(* IEC 61131-3 sources: stdmachine/plc/src/01_Types, 123 files *)

(* ---- E_ActStatus.st ---- *)
// Statut de l'action d'un objet (docs/04 § 5)
{attribute 'qualified_only'}
{attribute 'strict'}
TYPE E_ActStatus :
(
    Idle := 0,
    Busy := 1,
    Done := 2,
    Error := 3
) USINT;
END_TYPE

(* ---- E_AlarmEvent.st ---- *)
// Événement d'alarme (docs/14 § 5)
{attribute 'qualified_only'}
{attribute 'strict'}
TYPE E_AlarmEvent :
(
    Raised := 0,
    Cleared := 1,
    Acked := 2,
    Repeated := 3,
    Closed := 4
) USINT;
END_TYPE

(* ---- E_AlarmState.st ---- *)
// État d'une alarme active (docs/14 § 5)
{attribute 'qualified_only'}
{attribute 'strict'}
TYPE E_AlarmState :
(
    ActiveUnacked := 0,
    ActiveAcked := 1,
    ClearedUnacked := 2
) USINT;
END_TYPE

(* ---- E_BindTarget.st ---- *)
// Cible d'une liaison de résultat ou d'un SetVar (docs/06 § 2)
{attribute 'qualified_only'}
{attribute 'strict'}
TYPE E_BindTarget :
(
    None := 0,
    Var := 1,
    PartData := 2,
    PartId := 3,
    Verdict := 4,
    PartRemoved := 5,
    MoverData := 6,
    Output := 7
) USINT;
END_TYPE

(* ---- E_CalibState.st ---- *)
// État d'une calibration (docs/05 § 10.1)
{attribute 'qualified_only'}
{attribute 'strict'}
TYPE E_CalibState :
(
    Never := 0,
    Valid := 1,
    Expired := 2,
    Failed := 3,
    Running := 4
) USINT;
END_TYPE

(* ---- E_Cmd.st ---- *)
// Commandes d'état (docs/02 § 8). DrainStart et DrainCancel ne concernent que la machine (docs/05 § 5.7) :
// FB_PackML les ignore, le séquenceur général les traite.
{attribute 'qualified_only'}
{attribute 'strict'}
TYPE E_Cmd :
(
    None := 0,
    Reset := 1,
    Start := 2,
    Stop := 3,
    Hold := 4,
    Abort := 5,
    Clear := 6,
    DrainStart := 7,
    DrainCancel := 8
) USINT;
END_TYPE

(* ---- E_CmdResult.st ---- *)
// Résultat d'une commande (docs/05 § 2, docs/06 § 6.1)
{attribute 'qualified_only'}
{attribute 'strict'}
TYPE E_CmdResult :
(
    None := 0,
    Accepted := 1,
    Rejected := 2
) USINT;
END_TYPE

(* ---- E_Cmp.st ---- *)
// Comparaison d'un terme de condition (docs/05 § 3.7)
{attribute 'qualified_only'}
{attribute 'strict'}
TYPE E_Cmp :
(
    Eq := 0,
    Ne := 1,
    Lt := 2,
    Le := 3,
    Gt := 4,
    Ge := 5,
    IsTrue := 6,
    IsFalse := 7
) USINT;
END_TYPE

(* ---- E_Combine.st ---- *)
// Combinaison des termes d'une condition (docs/05 § 3.7)
{attribute 'qualified_only'}
{attribute 'strict'}
TYPE E_Combine :
(
    All := 0,
    Any := 1
) USINT;
END_TYPE

(* ---- E_CtxStatus.st ---- *)
// Statut d'un contexte d'exécution (docs/05 § 3.1)
{attribute 'qualified_only'}
{attribute 'strict'}
TYPE E_CtxStatus :
(
    Free := 0,
    Running := 1,
    WaitAction := 2,
    WaitCond := 3,
    WaitTime := 4,
    WaitJoin := 5,
    WaitStep := 6,
    Holding := 7,
    Done := 8,
    Failed := 9
) USINT;
END_TYPE

(* ---- E_DeclaredState.st ---- *)
// État déclaré de la machine (docs/12 § 2)
{attribute 'qualified_only'}
{attribute 'strict'}
TYPE E_DeclaredState :
(
    None := 0,
    PlannedStop := 1,
    Changeover := 2,
    WaitUpstream := 3,
    WaitDownstream := 4,
    PlannedMaintenance := 5,
    CorrectiveMaintenance := 6,
    Trials := 7,
    Cleaning := 8
) USINT;
END_TYPE

(* ---- E_DeployCmd.st ---- *)
// Commande de déploiement (docs/05 § 10)
{attribute 'qualified_only'}
{attribute 'strict'}
TYPE E_DeployCmd :
(
    None := 0,
    Verify := 1,
    Activate := 2,
    Cancel := 3
) USINT;
END_TYPE

(* ---- E_FailPolicy.st ---- *)
// Politique d'échec d'une instruction Action (docs/05 § 3.6)
{attribute 'qualified_only'}
{attribute 'strict'}
TYPE E_FailPolicy :
(
    StopStation := 0,
    Retry := 1,
    PartBad := 2,
    Goto := 3,
    Ignore := 4
) USINT;
END_TYPE

(* ---- E_ForceKind.st ---- *)
// Nature d'un forçage (docs/12 § 7)
{attribute 'qualified_only'}
{attribute 'strict'}
TYPE E_ForceKind :
(
    None := 0,
    DeclaredState := 1,
    StationOutOfProduction := 2,
    MoverOutOfService := 3
) USINT;
END_TYPE

(* ---- E_GroupRole.st ---- *)
// Rôle d'une fonction (docs/06 § 4)
{attribute 'qualified_only'}
{attribute 'strict'}
TYPE E_GroupRole :
(
    Entry := 0,
    Work := 1,
    Exit := 2,
    Reject := 3
) USINT;
END_TYPE

(* ---- E_Judgement.st ---- *)
// Jugement d'un résultat (docs/04 § 5)
{attribute 'qualified_only'}
{attribute 'strict'}
TYPE E_Judgement :
(
    None := 0,
    Ok := 1,
    Nok := 2,
    High := 3,
    Low := 4
) USINT;
END_TYPE

(* ---- E_ManualKind.st ---- *)
// Nature d'une demande du canal manuel (docs/05 § 7)
{attribute 'qualified_only'}
{attribute 'strict'}
TYPE E_ManualKind :
(
    Action := 0,
    JogStart := 1,
    JogStop := 2,
    Ack := 3,
    TeachPosition := 4
) USINT;
END_TYPE

(* ---- E_Mode.st ---- *)
// Modes de la machine (docs/02 § 8)
{attribute 'qualified_only'}
{attribute 'strict'}
TYPE E_Mode :
(
    Production := 0,
    Maintenance := 1
) USINT;
END_TYPE

(* ---- E_MoverState.st ---- *)
// État d'un mover dans le séquenceur général (docs/05 § 5.3)
{attribute 'qualified_only'}
{attribute 'strict'}
TYPE E_MoverState :
(
    Unknown := 0,
    Ready := 1,
    Routing := 2,
    Queued := 3,
    AtStation := 4,
    Buffered := 5,
    ToEmpty := 6,
    Error := 7,
    Halted := 8,
    OutOfService := 9
) USINT;
END_TYPE

(* ---- E_MoverVarReset.st ---- *)
// Règle de remise à zéro d'une variable de mover (docs/05 § 5.8)
{attribute 'qualified_only'}
{attribute 'strict'}
TYPE E_MoverVarReset :
(
    Never := 0,
    OnDeploy := 1,
    OnEmpty := 2
) USINT;
END_TYPE

(* ---- E_ObjState.st ---- *)
// États d'un objet (docs/04 § 5 et § 7.1)
{attribute 'qualified_only'}
{attribute 'strict'}
TYPE E_ObjState :
(
    NotInitialized := 0,
    Ready := 1,
    Busy := 2,
    Error := 3,
    Disabled := 4
) USINT;
END_TYPE

(* ---- E_Op.st ---- *)
// Jeu d'instructions (docs/06 § 2) ; version 2 du jeu : 17 à 23
{attribute 'qualified_only'}
{attribute 'strict'}
TYPE E_Op :
(
    Nop := 0,
    Action := 1,
    WaitCond := 2,
    WaitTime := 3,
    Jump := 4,
    JumpIfFalse := 5,
    Fork := 6,
    Join := 7,
    LoopInit := 8,
    LoopNext := 9,
    Call := 10,
    Return := 11,
    SetVar := 12,
    Alarm := 13,
    End := 14,
    StepBegin := 15,
    StepEnd := 16,
    WaitMover := 17,
    Prompt := 18,
    SavePos := 19,
    Route := 20,
    CalibStation := 21,
    ResetMoverVars := 22,
    SetOut := 23
) UINT;
END_TYPE

(* ---- E_OpStatus.st ---- *)
// Réponse d'une station à une demande d'opération (docs/05 § 4.1)
{attribute 'qualified_only'}
{attribute 'strict'}
TYPE E_OpStatus :
(
    Idle := 0,
    Running := 1,
    Done := 2,
    Failed := 3,
    Aborted := 4,
    Preparing := 5
) USINT;
END_TYPE

(* ---- E_OrderCmd.st ---- *)
// Commande d'OF (docs/05 § 5.6)
{attribute 'qualified_only'}
{attribute 'strict'}
TYPE E_OrderCmd :
(
    None := 0,
    Activate := 1,
    Suspend := 2,
    Cancel := 3
) USINT;
END_TYPE

(* ---- E_OrderState.st ---- *)
// État d'un OF dans la table du PLC (docs/05 § 5.6)
{attribute 'qualified_only'}
{attribute 'strict'}
TYPE E_OrderState :
(
    Free := 0,
    Active := 1,
    Suspended := 2,
    Done := 3
) USINT;
END_TYPE

(* ---- E_ParamKind.st ---- *)
// Nature d'un paramètre d'action résolu (docs/04 § 5)
{attribute 'qualified_only'}
{attribute 'strict'}
TYPE E_ParamKind :
(
    Unused := 0,
    Real := 1,
    Position := 2,
    SpeedIndex := 3,
    SpeedPercent := 4,
    Text := 5
) USINT;
END_TYPE

(* ---- E_PartStatus.st ---- *)
// État d'une pièce (docs/05 § 9)
{attribute 'qualified_only'}
{attribute 'strict'}
TYPE E_PartStatus :
(
    None := 0,
    InProcess := 1,
    Good := 2,
    Bad := 3,
    Exited := 4,
    Rejected := 5,
    Removed := 6
) USINT;
END_TYPE

(* ---- E_PlanarPosKind.st ---- *)
// Nature d'une position planaire (docs/05 § 6.1)
{attribute 'qualified_only'}
{attribute 'strict'}
TYPE E_PlanarPosKind :
(
    Work := 0,
    Queue := 1,
    Buffer := 2,
    Park := 3
) USINT;
END_TYPE

(* ---- E_QualityCmd.st ---- *)
// Commande de la surveillance des rebuts (docs/10 § 10)
{attribute 'qualified_only'}
{attribute 'strict'}
TYPE E_QualityCmd :
(
    None := 0,
    Release := 1,
    Reset := 2
) USINT;
END_TYPE

(* ---- E_QualityLevel.st ---- *)
// Niveau d'une portée qualité (docs/10 § 9)
{attribute 'qualified_only'}
{attribute 'strict'}
TYPE E_QualityLevel :
(
    Normal := 0,
    Warning := 1,
    Action := 2,
    Probation := 3
) USINT;
END_TYPE

(* ---- E_QualityReaction.st ---- *)
// Réaction de la surveillance des rebuts (docs/10 § 9)
{attribute 'qualified_only'}
{attribute 'strict'}
TYPE E_QualityReaction :
(
    WarnOnly := 0,
    StationHold := 1,
    MoverOut := 2,
    StopLoading := 3,
    MachineStop := 4
) USINT;
END_TYPE

(* ---- E_QualityScope.st ---- *)
// Portée de la surveillance des rebuts (docs/10 § 9)
{attribute 'qualified_only'}
{attribute 'strict'}
TYPE E_QualityScope :
(
    Station := 0,
    StationImputed := 1,
    Group := 2,
    Mover := 3,
    Machine := 4,
    Order := 5
) USINT;
END_TYPE

(* ---- E_RejectReason.st ---- *)
// Motif d'un refus de commande, traduit par la HMI (docs/06 § 6.1)
{attribute 'qualified_only'}
{attribute 'strict'}
TYPE E_RejectReason :
(
    None := 0,
    WrongState := 1,          // la commande n'est pas acceptée dans l'état courant
    StartBlocked := 2,        // état déclaré bloquant (docs/12 § 2)
    WrongMode := 3,           // mode Production / Maintenance
    NotAllowed := 4,          // station non réintégrable, cible inconnue
    Busy := 5,                // une opération ou une commande est en cours
    NotConfigured := 6,       // élément absent du déploiement
    TableFull := 7,           // table d'OF pleine
    PartsInProcess := 8,      // annulation d'un OF qui a encore des pièces
    Incompatible := 9         // projet plus récent que la bibliothèque (docs/02 § 7.3)
) USINT;
END_TYPE

(* ---- E_RetainedKind.st ---- *)
// Nature d'une valeur rémanente sauvegardée par la HMI (docs/02 § 7.4)
{attribute 'qualified_only'}
{attribute 'strict'}
TYPE E_RetainedKind :
(
    None := 0,
    StationVar := 1,       // variable persistante (calibration)
    MoverVar := 2,         // variable de mover
    ObjectCounters := 3,   // compteurs de maintenance d'un objet
    PlantCounters := 4,    // compteurs de production et de temps
    Calibration := 5       // état et date d'une calibration
) USINT;
END_TYPE

(* ---- E_Severity.st ---- *)
// Gravité d'une alarme (docs/04 § 5, docs/14 § 4)
{attribute 'qualified_only'}
{attribute 'strict'}
TYPE E_Severity :
(
    Info := 0,
    Warning := 1,
    StationFault := 2,
    MachineFault := 3,
    Quality := 4
) USINT;
END_TYPE

(* ---- E_SignalKind.st ---- *)
// Nature d'un signal de l'image E/S (docs/04 § 5)
{attribute 'qualified_only'}
{attribute 'strict'}
TYPE E_SignalKind :
(
    None := 0,
    DI := 1,
    DO := 2,
    AI := 3,
    AO := 4
) USINT;
END_TYPE

(* ---- E_StartResult.st ---- *)
// Réponse de I_Object.Start (docs/04 § 5)
{attribute 'qualified_only'}
{attribute 'strict'}
TYPE E_StartResult :
(
    Accepted := 0,
    Busy := 1,
    NotReady := 2,
    UnknownAction := 3,
    BadParam := 4,
    Interlocked := 5,
    Disabled := 6,
    ManualOnly := 7,
    NotConfigured := 8
) USINT;
END_TYPE

(* ---- E_State.st ---- *)
// États PackML réduits (docs/02 § 8, docs/05 § 2)
{attribute 'qualified_only'}
{attribute 'strict'}
TYPE E_State :
(
    Stopped := 0,
    Resetting := 1,
    Idle := 2,
    Execute := 3,
    Held := 4,
    Stopping := 5,
    Aborted := 6,
    Clearing := 7
) USINT;
END_TYPE

(* ---- E_StepGranularity.st ---- *)
// Granularité du pas à pas (docs/05 § 8)
{attribute 'qualified_only'}
{attribute 'strict'}
TYPE E_StepGranularity :
(
    Operation := 0,
    Step := 1,
    Action := 2
) USINT;
END_TYPE

(* ---- E_StopReason.st ---- *)
// Raison du dernier arrêt de la machine (docs/05 § 5.2, docs/14 § 4) : la cause système quand aucune alarme
// ne l'explique. Publiée dans ST_MachineStatus pour la HMI (toasts « OF terminé », « Machine vidée ») (D94)
{attribute 'qualified_only'}
{attribute 'strict'}
TYPE E_StopReason :
(
    None := 0,
    Alarm := 1,             // première alarme cause : nStopCauseGlobalId, nStopCauseCode
    Operator := 2,
    OrderComplete := 3,
    Drained := 4,
    Quality := 5
) USINT;
END_TYPE

(* ---- E_SystemVar.st ---- *)
// Variables système lues par la source System (docs/05 § 3.4)
{attribute 'qualified_only'}
{attribute 'strict'}
TYPE E_SystemVar :
(
    MoverPresent := 1,
    Slot := 2,
    OrderNo := 3,
    CycleCount := 4,
    LastCycleMs := 5
) INT;
END_TYPE

(* ---- E_TableKind.st ---- *)
// Nature d'une table (docs/06 § 2)
{attribute 'qualified_only'}
{attribute 'strict'}
TYPE E_TableKind :
(
    Operation := 0,
    Background := 1,
    Init := 2,
    Stop := 3,
    Clear := 4,
    Sub := 5,
    Calibration := 6,
    General := 10,
    GeneralSub := 11,
    MachineCalibration := 12
) USINT;
END_TYPE

(* ---- E_ValueSource.st ---- *)
// Source d'une valeur dans une instruction (docs/06 § 2)
{attribute 'qualified_only'}
{attribute 'strict'}
TYPE E_ValueSource :
(
    None := 0,
    Const := 1,
    Var := 2,
    PartData := 3,
    OpParam := 4,
    NamedPos := 5,
    Speed := 6,
    Text := 7,
    ObjValue := 8,
    System := 9,
    MoverData := 10,
    OrderParam := 11
) USINT;
END_TYPE

(* ---- E_VarType.st ---- *)
// Type d'une variable (docs/06 § 2)
{attribute 'qualified_only'}
{attribute 'strict'}
TYPE E_VarType :
(
    Number := 0,
    Bool := 1,
    Position := 2
) USINT;
END_TYPE

(* ---- E_Verdict.st ---- *)
// Verdict d'une pièce, donnée de pièce n° 1 (docs/05 § 9)
{attribute 'qualified_only'}
{attribute 'strict'}
TYPE E_Verdict :
(
    Undefined := 0,
    Good := 1,
    Bad := 2
) USINT;
END_TYPE

(* ---- E_WaitReason.st ---- *)
// Motif d'attente d'un mover en tampon (docs/05 § 5.4, 5.6, 5.7, docs/10)
{attribute 'qualified_only'}
{attribute 'strict'}
TYPE E_WaitReason :
(
    None := 0,
    NoStation := 1,
    OrderComplete := 2,
    NoOrder := 3,
    QualityStop := 4,
    Drain := 5,
    Held := 6
) USINT;
END_TYPE

(* ---- ST_ActParams.st ---- *)
// Paramètres résolus d'une action (docs/04 § 5)
{attribute 'pack_mode' := '1'}
TYPE ST_ActParams :
STRUCT
    aKind : ARRAY[1..GVL_Const.MAX_PARAMS] OF E_ParamKind;
    aReal : ARRAY[1..GVL_Const.MAX_PARAMS] OF LREAL;   // valeur, ou n° de vitesse, ou % de vitesse
    stPos : ST_Position;                               // le paramètre de type Position (un au plus)
    sText : STRING(80);                                // le paramètre de type Text (un au plus)
    nTimeoutMs : UDINT;                                // 0 = celui de la configuration ou du catalogue
END_STRUCT
END_TYPE

(* ---- ST_ActResults.st ---- *)
// Résultats d'une action (docs/04 § 5)
{attribute 'pack_mode' := '1'}
TYPE ST_ActResults :
STRUCT
    nCount : USINT;
    aReal : ARRAY[1..GVL_Const.MAX_PARAMS] OF LREAL;
    aJudgement : ARRAY[1..GVL_Const.MAX_PARAMS] OF E_Judgement;
    stPos : ST_Position;        // le résultat de type Position, s'il y en a un
    nPosIndex : USINT;          // rang du résultat de type Position, 0 = aucun
    sText : STRING(80);         // le résultat de type Text, s'il y en a un
    nTextIndex : USINT;         // rang du résultat de type Text, 0 = aucun
END_STRUCT
END_TYPE

(* ---- ST_AlarmAckRequest.st ---- *)
// Acquitter un avertissement (docs/06 § 6.2) ; nGlobalId 0 = tous les avertissements
{attribute 'pack_mode' := '1'}
TYPE ST_AlarmAckRequest :
STRUCT
    nSeq : UDINT;
    nGlobalId : UDINT;
    nCode : UINT;
    sUser : STRING(24);
END_STRUCT
END_TYPE

(* ---- ST_AlarmBuffer.st ---- *)
// Alarmes actives et tampon d'événements (docs/06 § 6.3)
{attribute 'pack_mode' := '1'}
TYPE ST_AlarmBuffer :
STRUCT
    nActive : UINT;
    aActive : ARRAY[1..GVL_Const.ALARM_ACTIVE] OF ST_AlarmEntry;
    nWriteSeq : UDINT;              // n° du dernier événement écrit
    aEvent : ARRAY[0..GVL_Const.ALARM_EVENTS - 1] OF ST_AlarmEventRec;
END_STRUCT
END_TYPE

(* ---- ST_AlarmContext.st ---- *)
// Contexte relevé à l'apparition d'une alarme (docs/14 § 5)
{attribute 'pack_mode' := '1'}
TYPE ST_AlarmContext :
STRUCT
    nTable : USINT;
    nStepId : UDINT;
    nMover : USINT;
    nSlot : USINT;
    sPartId : STRING(40);
    nAction : UINT;
END_STRUCT
END_TYPE

(* ---- ST_AlarmEntry.st ---- *)
// Alarme active (docs/04 § 10, docs/14)
{attribute 'pack_mode' := '1'}
TYPE ST_AlarmEntry :
STRUCT
    nGlobalId : UDINT;              // source : station × 1000 + n° local
    nCode : UINT;
    nSubCode : UDINT;
    eSeverity : E_Severity;
    eState : E_AlarmState;
    tRaised : LINT;
    tCleared : LINT;
    nRepeat : UINT;
    bCause : BOOL;                  // cause première d'un arrêt
    stCtx : ST_AlarmContext;
END_STRUCT
END_TYPE

(* ---- ST_AlarmEventRec.st ---- *)
// Événement d'alarme du tampon circulaire (docs/14 § 5)
{attribute 'pack_mode' := '1'}
TYPE ST_AlarmEventRec :
STRUCT
    nSeq : UDINT;
    eEvent : E_AlarmEvent;
    tTime : LINT;
    stAlarm : ST_AlarmEntry;
    sUser : STRING(24);
END_STRUCT
END_TYPE

(* ---- ST_Bind.st ---- *)
// Liaison d'un résultat (docs/06 § 2)
{attribute 'pack_mode' := '1'}
TYPE ST_Bind :
STRUCT
    eTarget : E_BindTarget;
    nIndex : INT;
END_STRUCT
END_TYPE

(* ---- ST_CalibDef.st ---- *)
// Déclaration d'une calibration d'une station (docs/05 § 10.1)
{attribute 'pack_mode' := '1'}
TYPE ST_CalibDef :
STRUCT
    nTable : USINT;             // table de type Calibration
    nId : UDINT;                // identifiant stable
    nValidityDays : UINT;       // 0 = n'expire jamais
END_STRUCT
END_TYPE

(* ---- ST_CalibStatus.st ---- *)
// État d'une calibration (docs/05 § 10.1)
{attribute 'pack_mode' := '1'}
TYPE ST_CalibStatus :
STRUCT
    nId : UDINT;
    eState : E_CalibState;
    tLast : LINT;
    sUser : STRING(24);
    nValidityDays : UINT;           // 0 = n'expire jamais
END_STRUCT
END_TYPE

(* ---- ST_CmdRequest.st ---- *)
// Commande d'état (docs/06 § 6.2) ; nTarget 0 = machine, 1..16 = station
{attribute 'pack_mode' := '1'}
TYPE ST_CmdRequest :
STRUCT
    nSeq : UDINT;
    nTarget : USINT;
    eCmd : E_Cmd;
    bSetMode : BOOL;                // changement de mode au lieu d'une commande
    eMode : E_Mode;
    sUser : STRING(24);
END_STRUCT
END_TYPE

(* ---- ST_CmdResponse.st ---- *)
// Réponse commune des handshakes (docs/06 § 6.1)
{attribute 'pack_mode' := '1'}
TYPE ST_CmdResponse :
STRUCT
    nSeq : UDINT;
    eResult : E_CmdResult;
    eReason : E_RejectReason;
    eState : E_State;               // état de la cible au moment de la réponse
    nDetail : UDINT;                // précision (n° d'élément, version demandée…)
END_STRUCT
END_TYPE

(* ---- ST_Condition.st ---- *)
// Condition (docs/05 § 3.7) ; une condition sans terme est vraie
{attribute 'pack_mode' := '1'}
TYPE ST_Condition :
STRUCT
    eCombine : E_Combine;
    nTerms : USINT;
    aTerm : ARRAY[1..GVL_Const.MAX_COND_TERMS] OF ST_CondTerm;
END_STRUCT
END_TYPE

(* ---- ST_CondTerm.st ---- *)
// Terme de condition (docs/05 § 3.7)
{attribute 'pack_mode' := '1'}
TYPE ST_CondTerm :
STRUCT
    stLeft : ST_Value;
    eCmp : E_Cmp;
    stRight : ST_Value;
END_STRUCT
END_TYPE

(* ---- ST_Context.st ---- *)
// Contexte d'exécution d'une station (docs/05 § 3.1)
TYPE ST_Context :
STRUCT
    eStatus : E_CtxStatus;
    nTable : USINT;                 // table en cours
    nPC : INT;                      // index d'instruction absolu dans aInstr
    aRetTable : ARRAY[1..GVL_Const.MAX_CALL_DEPTH] OF USINT;
    aRetPC : ARRAY[1..GVL_Const.MAX_CALL_DEPTH] OF INT;
    nDepth : USINT;
    nParent : USINT;                // contexte qui a fait le Fork, 0 sinon
    nForkPC : INT;                  // Fork de rattachement
    nChildren : USINT;              // branches filles encore actives
    bBranchFailed : BOOL;           // une branche a terminé l'opération (pièce mauvaise)
    nRetry : USINT;
    fWaitMs : LREAL;
    nStepId : UDINT;                // carte en cours
    nStepDepth : USINT;
    nErrorCode : UINT;
    bStarted : BOOL;                // l'instruction courante a déjà été lancée (Action, Prompt…)
    bStepReleased : BOOL;           // pas à pas : point d'arrêt déjà franchi pour cette instruction
END_STRUCT
END_TYPE

(* ---- ST_CtxStatus.st ---- *)
// Statut publié d'un contexte (docs/05 § 4.5)
{attribute 'pack_mode' := '1'}
TYPE ST_CtxStatus :
STRUCT
    eStatus : E_CtxStatus;
    nTable : USINT;
    nPC : INT;
    nStepId : UDINT;
    nNextStepId : UDINT;
    nObject : UINT;
    nAction : UINT;
    nRetry : USINT;
    fWaitMs : REAL;
    stNextParams : ST_ActParams;    // pas à pas : paramètres résolus de la prochaine action
END_STRUCT
END_TYPE

(* ---- ST_DeployError.st ---- *)
// Erreur rendue par le chargeur (docs/05 § 10)
{attribute 'pack_mode' := '1'}
TYPE ST_DeployError :
STRUCT
    nCode : UINT;                   // voir FB_Loader
    nStation : USINT;               // 0 = machine
    nTable : USINT;
    nInstr : INT;
    nObject : UINT;
    nDetail : UDINT;
END_STRUCT
END_TYPE

(* ---- ST_DeployRequest.st ---- *)
// Vérifier, activer ou annuler la zone d'attente (docs/05 § 10)
{attribute 'pack_mode' := '1'}
TYPE ST_DeployRequest :
STRUCT
    nSeq : UDINT;
    eCmd : E_DeployCmd;
    nCrcMachine : UDINT;
    aCrcStation : ARRAY[1..GVL_Const.MAX_STATIONS] OF UDINT;
    nCrcRecipes : UDINT;
    nInstrSetRequired : UINT;       // docs/02 § 7.3
    nCatalogRequired : UINT;
    sUser : STRING(24);
END_STRUCT
END_TYPE

(* ---- ST_DeployResponse.st ---- *)
// Réponse du chargeur (docs/05 § 10)
{attribute 'pack_mode' := '1'}
TYPE ST_DeployResponse :
STRUCT
    nSeq : UDINT;
    eResult : E_CmdResult;
    nErrors : USINT;
    aError : ARRAY[1..32] OF ST_DeployError;
END_STRUCT
END_TYPE

(* ---- ST_ForceCommand.st ---- *)
// Poser ou lever un forçage (docs/12 § 7)
{attribute 'pack_mode' := '1'}
TYPE ST_ForceCommand :
STRUCT
    nSeq : UDINT;
    eKind : E_ForceKind;
    bSet : BOOL;                    // faux = lever
    nTarget : USINT;                // station ou mover
    eDeclared : E_DeclaredState;
    bStartBlocked : BOOL;
    bImmediate : BOOL;              // mover hors service immédiatement
    nReason : USINT;                // code de motif
    tUntil : LINT;                  // échéance, 0 = aucune (gérée par la HMI)
    sUser : STRING(24);
END_STRUCT
END_TYPE

(* ---- ST_GroupCfg.st ---- *)
// Fonction (docs/06 § 4)
{attribute 'pack_mode' := '1'}
TYPE ST_GroupCfg :
STRUCT
    bUsed : BOOL;
    sName : STRING(40);
    eRole : E_GroupRole;
    nStationMask : UINT;        // bit n-1 = station n
    nOperations : USINT;
    nPriority : USINT;          // 1..9
END_STRUCT
END_TYPE

(* ---- ST_Instr.st ---- *)
// Instruction (docs/06 § 2), 154 octets
{attribute 'pack_mode' := '1'}
TYPE ST_Instr :
STRUCT
    eOp : E_Op;
    nStepId : UDINT;            // carte de l'éditeur ; 0 = instruction technique
    nObject : UINT;             // Action : n° local de l'objet
    nAction : UINT;             // Action : n° d'action du catalogue
    aParam : ARRAY[1..GVL_Const.MAX_PARAMS] OF ST_Value;
    aBind : ARRAY[1..GVL_Const.MAX_PARAMS] OF ST_Bind;
    aArg : ARRAY[1..GVL_Const.MAX_ARGS] OF DINT;
    nTimeoutMs : UDINT;         // 0 = défaut (configuration de l'objet, puis catalogue)
    eOnFail : E_FailPolicy;
    nRetries : USINT;
    nFailTarget : INT;          // Goto : index d'instruction
END_STRUCT
END_TYPE

(* ---- ST_Interlock.st ---- *)
// Verrouillage (docs/06 § 2)
{attribute 'pack_mode' := '1'}
TYPE ST_Interlock :
STRUCT
    nObject : UINT;             // objet protégé
    nActionMask : UDINT;        // bit n-1 = action n ; 0 = toutes les actions de mouvement
    nCond : INT;                // condition qui doit rester vraie
END_STRUCT
END_TYPE

(* ---- ST_LaunchRequest.st ---- *)
// Maintenance : lancer une table d'une station (docs/06 § 6.2)
{attribute 'pack_mode' := '1'}
TYPE ST_LaunchRequest :
STRUCT
    nSeq : UDINT;
    nStation : USINT;               // 0 = calibration machine
    nTable : USINT;
    nMover : USINT;                 // 0 = sans mover
    nSlot : USINT;
    aParam : ARRAY[1..GVL_Const.MAX_PARAMS] OF LREAL;
    sUser : STRING(24);
END_STRUCT
END_TYPE

(* ---- ST_MachineData.st ---- *)
// Configuration machine déployée (docs/06 § 4)
{attribute 'pack_mode' := '1'}
TYPE ST_MachineData :
STRUCT
    sMachineName : STRING(40);
    sProjectId : STRING(40);
    sProjectHash : STRING(64);
    tDeployed : LINT;
    sDeployedBy : STRING(40);
    nMovers : USINT;
    nSlots : USINT;
    fOverride : LREAL;
    nRejectGroup : USINT;       // 0 = aucune fonction de rebut
    nNoStationMs : UDINT;       // délai avant « mover à vider »
    nMoverVar : USINT;
    aMoverVar : ARRAY[1..GVL_Const.MAX_MOVER_VARS] OF ST_MoverVarDef;
    aGroup : ARRAY[1..GVL_Const.MAX_GROUPS] OF ST_GroupCfg;
    aStation : ARRAY[1..GVL_Const.MAX_STATIONS] OF ST_StationCfg;
    nPlanarPos : INT;
    aPlanarPos : ARRAY[1..GVL_Const.MAX_PLANAR_POS] OF ST_PlanarPos;
    nParkPos : INT;
    nMachineObj : UINT;
    aMachineObj : ARRAY[1..GVL_Const.MAX_MACHINE_OBJ] OF ST_ObjConfig;
    aTable : ARRAY[1..GVL_Const.MAX_TABLES] OF ST_TableDir;
    nInstrCount : INT;
    aInstr : ARRAY[1..GVL_Const.MAX_INSTR] OF ST_Instr;
    aCond : ARRAY[1..GVL_Const.MAX_COND] OF ST_Condition;
    aText : ARRAY[1..GVL_Const.MAX_TEXTS] OF STRING(80);
    stQuality : ST_QualityCfg;
    nCalibCount : USINT;
    aCalib : ARRAY[1..GVL_Const.CALIB_PER_STATION] OF ST_CalibDef;  // calibrations machine
END_STRUCT
END_TYPE

(* ---- ST_MachineForce.st ---- *)
// Forçages actifs (docs/12 § 7), persistants
{attribute 'pack_mode' := '1'}
TYPE ST_MachineForce :
STRUCT
    eDeclared : E_DeclaredState;
    bStartBlocked : BOOL;
    nReason : USINT;
    tSince : LINT;
    tUntil : LINT;
    sBy : STRING(24);
    aStation : ARRAY[1..GVL_Const.MAX_STATIONS] OF ST_StationForce;
    aMover : ARRAY[1..GVL_Const.MAX_MOVERS] OF ST_MoverForce;
END_STRUCT
END_TYPE

(* ---- ST_MachineStatus.st ---- *)
// Statut de la machine (docs/06 § 6.3)
{attribute 'pack_mode' := '1'}
TYPE ST_MachineStatus :
STRUCT
    eState : E_State;
    eMode : E_Mode;
    fEffOverride : REAL;
    nBeacon : UINT;
    bFault : BOOL;
    tStateSince : LINT;
    nStopCauseGlobalId : UDINT;     // cause première (docs/14 § 4)
    nStopCauseCode : UINT;
    eStopReason : E_StopReason;     // D94
    nActiveOrder : UDINT;           // n° interne, 0 = aucun
    aOrder : ARRAY[1..GVL_Const.MAX_ORDERS] OF ST_OrderState;
    bDrain : BOOL;                  // fin des pièces en cours (docs/05 § 5.7)
    nPartsInProcess : UINT;
    bLoadingLocked : BOOL;          // arrêt du chargement qualité
    eDeclared : E_DeclaredState;
    bStartBlocked : BOOL;
    tPlcClock : LINT;               // UTC
    nPlcHeartbeat : UDINT;
    sProjectHash : STRING(64);
    tDeployed : LINT;
    nCalib : USINT;
    aCalib : ARRAY[1..GVL_Const.CALIB_PER_STATION] OF ST_CalibStatus;
    stPrompt : ST_PromptState;      // calibration machine
    bHmiLost : BOOL;                // battement de la HMI perdu (alarme 917)
END_STRUCT
END_TYPE

(* ---- ST_ManualRequest.st ---- *)
// Demande du canal manuel (docs/05 § 7)
{attribute 'pack_mode' := '1'}
TYPE ST_ManualRequest :
STRUCT
    nSeq : UDINT;
    eKind : E_ManualKind;
    nObject : UINT;                 // n° local
    nAction : UINT;
    stParams : ST_ActParams;        // résolus par la HMI
    nTeachPos : INT;                // position nommée à apprendre
    nTeachMask : USINT;             // bits X, Y, Z, C
    aTeachFrom : ARRAY[1..4] OF UINT;   // objets qui fournissent X, Y, Z, C
    sUser : STRING(24);
END_STRUCT
END_TYPE

(* ---- ST_ManualResponse.st ---- *)
// Réponse du canal manuel (docs/05 § 7)
{attribute 'pack_mode' := '1'}
TYPE ST_ManualResponse :
STRUCT
    nSeq : UDINT;
    eResult : E_CmdResult;
    eReason : E_RejectReason;
    eStart : E_StartResult;
    eActStatus : E_ActStatus;
    nErrorCode : UINT;
    nSubCode : UDINT;
    stResults : ST_ActResults;
    stTaught : ST_Position;
END_STRUCT
END_TYPE

(* ---- ST_MoverCtx.st ---- *)
// Contexte d'un mover dans le séquenceur général (docs/05 § 5.3)
TYPE ST_MoverCtx :
STRUCT
    eState : E_MoverState;
    eWait : E_WaitReason;
    nTable : INT;
    nPC : INT;
    aRetTable : ARRAY[1..GVL_Const.MAX_CALL_DEPTH] OF INT;
    aRetPC : ARRAY[1..GVL_Const.MAX_CALL_DEPTH] OF INT;
    nDepth : USINT;
    nTargetGroup : USINT;
    nTargetOp : USINT;
    nTargetSlot : USINT;
    aOpParam : ARRAY[1..GVL_Const.MAX_PARAMS] OF LREAL;   // paramètres résolus à l'émission de Route
    nStation : USINT;               // station réservée ou occupée, 0 = aucune
    nDest : INT;                    // position planaire de destination
    nPos : INT;                     // position planaire occupée, 0 = entre deux positions
    nReqId : UDINT;
    bRequestPosted : BOOL;
    nRouteRetry : UDINT;
    tWaitStart : LINT;
    fWaitMs : LREAL;
    fMoveMs : LREAL;                // durée du déplacement en cours
    fStillMs : LREAL;               // à l'arrêt dans la fenêtre d'arrivée
    bQualityLock : BOOL;
    bOutOfService : BOOL;
    bImmediate : BOOL;
    bAbsent : BOOL;                 // hors service et absent du plan (D85)
    bStationAborted : BOOL;         // la station de l'opération est passée Aborted (docs/05 § 6.4)
    bToEmptyPark : BOOL;            // en route vers le parcage pour être vidé
    aBadAtArrival : ARRAY[1..GVL_Const.MAX_SLOTS] OF BOOL;     // verdict déjà mauvais à l'arrivée (docs/10 § 9)
    aDefectBad : ARRAY[1..GVL_Const.MAX_SLOTS] OF BOOL;        // mauvaise sur défaut de station (docs/10 § 2)
    aHidden : ARRAY[1..8] OF LREAL; // compteurs de boucle du process général (D93)
    tOpStart : LINT;                // début de l'opération en cours
    fX : LREAL;                     // position actuelle sur le plan
    fY : LREAL;
    fC : LREAL;
    aSlot : ARRAY[1..GVL_Const.MAX_SLOTS] OF ST_Part;
    aVar : ARRAY[1..GVL_Const.MAX_MOVER_VARS] OF LREAL;          // variables de mover (docs/05 § 5.8)
    aVarPos : ARRAY[1..GVL_Const.MAX_MOVER_VARS] OF ST_Position;
    aVarId : ARRAY[1..GVL_Const.MAX_MOVER_VARS] OF UDINT;
END_STRUCT
END_TYPE

(* ---- ST_MoverForce.st ---- *)
// Forçage d'un mover (docs/12 § 4)
{attribute 'pack_mode' := '1'}
TYPE ST_MoverForce :
STRUCT
    bOutOfService : BOOL;
    bImmediate : BOOL;
    nReason : USINT;
    tSince : LINT;
    sBy : STRING(24);
END_STRUCT
END_TYPE

(* ---- ST_MoverStatus.st ---- *)
// Statut d'un mover (docs/06 § 6.3)
{attribute 'pack_mode' := '1'}
TYPE ST_MoverStatus :
STRUCT
    eState : E_MoverState;
    eWait : E_WaitReason;
    fX : REAL;
    fY : REAL;
    fC : REAL;
    nStation : USINT;
    nDest : INT;
    nTargetGroup : USINT;
    nTable : INT;
    nPC : INT;
    nStepId : UDINT;
    bOutOfService : BOOL;
    bQualityLock : BOOL;
    bAbsent : BOOL;
    aSlot : ARRAY[1..GVL_Const.MAX_SLOTS] OF ST_SlotStatus;
    aVar : ARRAY[1..GVL_Const.MAX_MOVER_VARS] OF LREAL;
    aVarPos : ARRAY[1..GVL_Const.MAX_MOVER_VARS] OF ST_Position;
    aVarId : ARRAY[1..GVL_Const.MAX_MOVER_VARS] OF UDINT;
END_STRUCT
END_TYPE

(* ---- ST_MoverVarDef.st ---- *)
// Déclaration d'une variable de mover (docs/05 § 5.8)
{attribute 'pack_mode' := '1'}
TYPE ST_MoverVarDef :
STRUCT
    nId : UDINT;                // identifiant stable
    sName : STRING(24);
    eType : E_VarType;
    sUnit : STRING(8);
    fInit : LREAL;
    stInitPos : ST_Position;
    eReset : E_MoverVarReset;
END_STRUCT
END_TYPE

(* ---- ST_MoverVarRequest.st ---- *)
// Écrire ou remettre à zéro une variable de mover (docs/05 § 5.8)
{attribute 'pack_mode' := '1'}
TYPE ST_MoverVarRequest :
STRUCT
    nSeq : UDINT;
    nMover : USINT;
    nVar : USINT;                   // rang
    bReset : BOOL;                  // valeur initiale
    fValue : LREAL;
    stPos : ST_Position;
    sUser : STRING(24);
END_STRUCT
END_TYPE

(* ---- ST_NamedPos.st ---- *)
// Position nommée (docs/06 § 2)
{attribute 'pack_mode' := '1'}
TYPE ST_NamedPos :
STRUCT
    stPos : ST_Position;
    fApproach : LREAL;
    bTaught : BOOL;
END_STRUCT
END_TYPE

(* ---- ST_ObjConfig.st ---- *)
// Configuration d'un objet, écrite par la HMI au déploiement (docs/04 § 5)
{attribute 'pack_mode' := '1'}
TYPE ST_ObjConfig :
STRUCT
    nType : UINT;
    nLocalId : UINT;
    nParentId : UINT;
    nStableId : UDINT;          // empreinte de l'identifiant de l'objet dans le projet (D92)
    sName : STRING(40);
    bSimulated : BOOL;
    bDisabled : BOOL;
    fOverride : LREAL;                                          // 0..100
    aSignal : ARRAY[1..GVL_Const.MAX_SIGNALS] OF ST_SignalRef;  // S1..S8
    nDevice : INT;                                              // D : élément de pool matériel, 0 = aucun
    aParam : ARRAY[1..GVL_Const.MAX_OBJ_PARAMS] OF LREAL;       // P1..P24
    aSpeedPct : ARRAY[1..GVL_Const.MAX_SPEEDS] OF LREAL;        // V1..V8, 0 = non défini
    aTimeoutMs : ARRAY[1..GVL_Const.MAX_ACTION_TIMEOUTS] OF UDINT; // par n° d'action, 0 = défaut du catalogue
END_STRUCT
END_TYPE

(* ---- ST_ObjectInfo.st ---- *)
// Identité d'un objet (docs/04 § 5)
{attribute 'pack_mode' := '1'}
TYPE ST_ObjectInfo :
STRUCT
    nGlobalId : UDINT;          // n° de station × 1000 + n° local (station 0 = machine)
    nStation : UINT;
    nLocalId : UINT;            // 1..64 dans la station
    nParentId : UINT;           // n° local du parent, 0 = la station
    nType : UINT;               // n° de type du catalogue
    nPoolIndex : UINT;
    nStableId : UDINT;          // identifiant stable donné par la HMI (D92)
    sName : STRING(40);
END_STRUCT
END_TYPE

(* ---- ST_ObjStatus.st ---- *)
// Statut d'un objet publié à chaque cycle (docs/04 § 5)
{attribute 'pack_mode' := '1'}
TYPE ST_ObjStatus :
STRUCT
    eState : E_ObjState;
    eActStatus : E_ActStatus;
    nAction : USINT;            // action en cours ou dernière action
    bManual : BOOL;
    nErrorCode : UINT;
    nSubCode : UDINT;
    fEffOverride : REAL;        // %
    bOverrideHalted : BOOL;     // mouvement suspendu par override à 0 %
    bSimulated : BOOL;
    nInterlock : USINT;         // verrouillage qui bloque, 0 = aucun
    fProgress : REAL;           // 0..1 avancement estimé, -1 = inconnu
    nElapsedMs : UDINT;
    nActionCount : UDINT;       // maintenance, persistant
    nErrorCount : UDINT;        // maintenance, persistant
    fMotionHours : REAL;        // maintenance, persistant
    nTimeoutMs : UDINT;         // timeout effectif estimé (affichage)
    aValue : ARRAY[1..GVL_Const.MAX_VALUES] OF LREAL;   // E1..E4
END_STRUCT
END_TYPE

(* ---- ST_OpMap.st ---- *)
// (fonction, opération) → table (docs/06 § 4)
{attribute 'pack_mode' := '1'}
TYPE ST_OpMap :
STRUCT
    nGroup : USINT;
    nOperationNo : USINT;       // 1..8
    nTable : USINT;
    bPrepare : BOOL;            // la table contient WaitMover (docs/05 § 4.1)
END_STRUCT
END_TYPE

(* ---- ST_OpRequest.st ---- *)
// Demande d'opération du séquenceur général à une station (docs/05 § 4.1)
TYPE ST_OpRequest :
STRUCT
    nReqId : UDINT;                 // change à chaque nouvelle demande
    nGroup : USINT;
    nOperation : USINT;
    nMover : USINT;
    nSlot : USINT;                  // 0 = tous
    bMoverAtStation : BOOL;         // préparation : faux tant que le mover n'est pas arrivé
    bCancel : BOOL;                 // préparation annulée (Stop)
    aParam : ARRAY[1..GVL_Const.MAX_PARAMS] OF LREAL;
END_STRUCT
END_TYPE

(* ---- ST_OpResponse.st ---- *)
// Réponse d'une station (docs/05 § 4.1)
TYPE ST_OpResponse :
STRUCT
    nReqId : UDINT;
    eStatus : E_OpStatus;
    nErrorCode : UINT;
    nOutMask : UINT;                // bit k-1 = sortie k définie
    aOut : ARRAY[1..GVL_Const.MAX_OUTPUTS] OF LREAL;
    stOutPos : ST_Position;
END_STRUCT
END_TYPE

(* ---- ST_OrderRequest.st ---- *)
// OF : activer, suspendre, annuler (docs/05 § 5.6)
{attribute 'pack_mode' := '1'}
TYPE ST_OrderRequest :
STRUCT
    nSeq : UDINT;
    eCmd : E_OrderCmd;
    nOrder : UDINT;                 // n° interne
    sNumber : STRING(40);
    sReference : STRING(40);
    nQuantity : UDINT;
    nGoodDone : UDINT;              // compteurs déjà faits (reprise)
    nBadDone : UDINT;
    aParam : ARRAY[1..GVL_Const.MAX_ORDER_PARAMS] OF LREAL;
    sUser : STRING(24);
END_STRUCT
END_TYPE

(* ---- ST_OrderState.st ---- *)
// OF dans la table du séquenceur général (docs/05 § 5.6)
{attribute 'pack_mode' := '1'}
TYPE ST_OrderState :
STRUCT
    nOrder : UDINT;                 // n° interne, 0 = libre
    eState : E_OrderState;
    sNumber : STRING(40);
    sReference : STRING(40);
    nQuantity : UDINT;
    nGood : UDINT;
    nBad : UDINT;
    nInProcess : UDINT;
    aParam : ARRAY[1..GVL_Const.MAX_ORDER_PARAMS] OF LREAL;
    stQuality : ST_QualityTrack;    // budget de rebuts de l'OF (docs/10 § 4.3)
END_STRUCT
END_TYPE

(* ---- ST_OverrideRequest.st ---- *)
// Override d'un nœud (docs/06 § 6.2) ; nStation 0 = machine ; nObject 0 = la station ou la machine
{attribute 'pack_mode' := '1'}
TYPE ST_OverrideRequest :
STRUCT
    nSeq : UDINT;
    nStation : USINT;
    nObject : UINT;
    fValue : LREAL;                 // 0..100 %
    bManual : BOOL;                 // override manuel de l'axe
    sUser : STRING(24);
END_STRUCT
END_TYPE

(* ---- ST_Part.st ---- *)
// Pièce portée par un emplacement de mover (docs/05 § 9)
{attribute 'pack_mode' := '1'}
TYPE ST_Part :
STRUCT
    bPresent : BOOL;
    sPartId : STRING(40);
    nOrder : UDINT;                 // n° interne de l'OF de la pièce
    eStatus : E_PartStatus;
    bBadHandled : BOOL;
    nOps : USINT;
    aOps : ARRAY[1..GVL_Const.MAX_PART_OPS] OF ST_PartOp;
    aData : ARRAY[1..GVL_Const.MAX_PART_DATA] OF LREAL;   // donnée 1 = verdict (0 non défini, 1 bon, 2 mauvais)
    tCreated : LINT;                // UTC, 100 ns depuis 1601
END_STRUCT
END_TYPE

(* ---- ST_PartOp.st ---- *)
// Opération subie par une pièce (docs/05 § 9)
{attribute 'pack_mode' := '1'}
TYPE ST_PartOp :
STRUCT
    nStation : USINT;
    nGroup : USINT;
    eVerdictAfter : E_Verdict;
END_STRUCT
END_TYPE

(* ---- ST_PartRequest.st ---- *)
// Confirmer le retrait des pièces d'un mover à vider (docs/06 § 6.2)
{attribute 'pack_mode' := '1'}
TYPE ST_PartRequest :
STRUCT
    nSeq : UDINT;
    nMover : USINT;
    sUser : STRING(24);
END_STRUCT
END_TYPE

(* ---- ST_PlanarPos.st ---- *)
// Position planaire (docs/05 § 6.1), toujours en frame 0
{attribute 'pack_mode' := '1'}
TYPE ST_PlanarPos :
STRUCT
    stPos : ST_Position;
    eKind : E_PlanarPosKind;
    nStation : USINT;
END_STRUCT
END_TYPE

(* ---- ST_PlcIdentity.st ---- *)
// Identité du PLC (docs/06 § 2) ; nInterfaceVersion est toujours le premier champ
{attribute 'pack_mode' := '1'}
TYPE ST_PlcIdentity :
STRUCT
    nInterfaceVersion : UINT;
    nInstrSetVersion : UINT;
    nCatalogVersion : UINT;
    sLibVersion : STRING(20);
    aPoolSize : ARRAY[1..149] OF UINT;  // par n° de type, 0 = type absent
    nRetainId : ULINT;
END_STRUCT
END_TYPE

(* ---- ST_Position.st ---- *)
// Toujours X, Y, Z, C + frame (docs/04 § 5). Le frame n'est exploité que par un robot Stäubli (D86).
{attribute 'pack_mode' := '1'}
TYPE ST_Position :
STRUCT
    fX : LREAL;                 // mm
    fY : LREAL;                 // mm
    fZ : LREAL;                 // mm
    fC : LREAL;                 // degrés
    nFrame : INT;               // 0 = repère machine ou repère des axes
END_STRUCT
END_TYPE

(* ---- ST_PressCurve.st ---- *)
// Courbe de presse (docs/05 § 9)
{attribute 'pack_mode' := '1'}
TYPE ST_PressCurve :
STRUCT
    nCurveId : UDINT;
    nPoints : UINT;
    aStroke : ARRAY[1..GVL_Const.CURVE_POINTS] OF REAL;
    aForce : ARRAY[1..GVL_Const.CURVE_POINTS] OF REAL;
END_STRUCT
END_TYPE

(* ---- ST_PressRecipe.st ---- *)
// Recette de presse (docs/06 § 4)
{attribute 'pack_mode' := '1'}
TYPE ST_PressRecipe :
STRUCT
    bUsed : BOOL;
    nStation : USINT;
    nObject : UINT;
    nRecipeNo : USINT;
    nSegments : USINT;
    aSeg : ARRAY[1..GVL_Const.MAX_PRESS_SEGMENTS] OF ST_PressSegment;
END_STRUCT
END_TYPE

(* ---- ST_PressSegment.st ---- *)
// Segment d'une recette de presse (docs/06 § 4)
{attribute 'pack_mode' := '1'}
TYPE ST_PressSegment :
STRUCT
    eTarget : USINT;            // 0 course, 1 force
    fTarget : LREAL;
    fSpeedPct : LREAL;
    fForceMin : LREAL;
    fForceMax : LREAL;
    fStrokeMin : LREAL;
    fStrokeMax : LREAL;
END_STRUCT
END_TYPE

(* ---- ST_PromptAnswer.st ---- *)
// Réponse de l'opérateur (docs/06 § 6.2) ; nStation 0 = calibration machine
{attribute 'pack_mode' := '1'}
TYPE ST_PromptAnswer :
STRUCT
    nSeq : UDINT;
    nStation : USINT;
    nPromptId : UDINT;
    bConfirm : BOOL;                // faux = annuler
    fValue : LREAL;
    sUser : STRING(24);
END_STRUCT
END_TYPE

(* ---- ST_PromptState.st ---- *)
// Demande à l'opérateur en cours (docs/05 § 10.1)
{attribute 'pack_mode' := '1'}
TYPE ST_PromptState :
STRUCT
    nPromptId : UDINT;              // 0 = aucune demande
    nText : INT;                    // n° de texte de la table
    bInput : BOOL;                  // saisie d'une valeur (sinon confirmation)
END_STRUCT
END_TYPE

(* ---- ST_QualityCfg.st ---- *)
// Configuration déployée de la surveillance des rebuts (docs/10 § 9)
{attribute 'pack_mode' := '1'}
TYPE ST_QualityCfg :
STRUCT
    aDefault : ARRAY[0..5] OF ST_QualityRule;                   // par E_QualityScope
    aStationRule : ARRAY[1..GVL_Const.MAX_STATIONS] OF ST_QualityRule;
    aStationInherits : ARRAY[1..GVL_Const.MAX_STATIONS] OF BOOL;
    aGroupRule : ARRAY[1..GVL_Const.MAX_GROUPS] OF ST_QualityRule;
    aGroupInherits : ARRAY[1..GVL_Const.MAX_GROUPS] OF BOOL;
    aGroupImpute : ARRAY[1..GVL_Const.MAX_GROUPS] OF UINT;      // masque des fonctions amont imputées, 0 = n'impute pas
    nOrderBudgetCount : UDINT;                                  // budget de rebuts d'OF en nombre, 0 = aucun
    fOrderBudgetPct : REAL;                                     // ou en %, 0 = aucun
END_STRUCT
END_TYPE

(* ---- ST_QualityCommand.st ---- *)
// Libérer ou remettre à zéro une portée qualité (docs/10 § 10)
{attribute 'pack_mode' := '1'}
TYPE ST_QualityCommand :
STRUCT
    nSeq : UDINT;
    eCmd : E_QualityCmd;
    eScope : E_QualityScope;
    nIndex : USINT;
    nReason : USINT;
    sUser : STRING(24);
END_STRUCT
END_TYPE

(* ---- ST_QualityRule.st ---- *)
// Réglage d'une portée qualité (docs/10 § 9)
{attribute 'pack_mode' := '1'}
TYPE ST_QualityRule :
STRUCT
    nConsecWarn : USINT;        // 0 = désactivé
    nConsecAction : USINT;
    nWindow : USINT;            // 1..255
    nMinSample : USINT;
    fRateWarn : REAL;           // %, 0 = désactivé
    fRateAction : REAL;
    eReactionConsec : E_QualityReaction;
    eReactionRate : E_QualityReaction;
END_STRUCT
END_TYPE

(* ---- ST_QualityStatus.st ---- *)
// État de la surveillance des rebuts (docs/10 § 9)
{attribute 'pack_mode' := '1'}
TYPE ST_QualityStatus :
STRUCT
    aStation : ARRAY[1..GVL_Const.MAX_STATIONS] OF ST_QualityTrack;
    aStationImputed : ARRAY[1..GVL_Const.MAX_STATIONS] OF ST_QualityTrack;
    aGroup : ARRAY[1..GVL_Const.MAX_GROUPS] OF ST_QualityTrack;
    aMover : ARRAY[1..GVL_Const.MAX_MOVERS] OF ST_QualityTrack;
    stMachine : ST_QualityTrack;
    bLoadingLocked : BOOL;
END_STRUCT
END_TYPE

(* ---- ST_QualityTrack.st ---- *)
// État d'une instance de portée qualité (docs/10 § 9)
{attribute 'pack_mode' := '1'}
TYPE ST_QualityTrack :
STRUCT
    nConsec : USINT;
    aWindow : ARRAY[0..31] OF BYTE;     // 256 résultats en bits (1 = mauvais)
    nHead : USINT;
    nCount : USINT;
    nBadInWindow : USINT;
    nProbationLeft : USINT;
    eLevel : E_QualityLevel;
    bLocked : BOOL;
    nTotalGood : UDINT;
    nTotalBad : UDINT;
END_STRUCT
END_TYPE

(* ---- ST_RestoreRequest.st ---- *)
// Restauration des valeurs rémanentes, par pages de 256 (docs/05 § 10, étape 6)
{attribute 'pack_mode' := '1'}
TYPE ST_RestoreRequest :
STRUCT
    nSeq : UDINT;
    nPage : UINT;                   // 0 = première page (efface la liste en cours)
    bLast : BOOL;                   // dernière page : appliquer
    nCount : UINT;
    aItem : ARRAY[1..256] OF ST_RetainedItem;
    sUser : STRING(24);
END_STRUCT
END_TYPE

(* ---- ST_RetainedItem.st ---- *)
// Valeur rémanente sauvegardée par la HMI, rangée par identifiant (docs/02 § 7.4)
{attribute 'pack_mode' := '1'}
TYPE ST_RetainedItem :
STRUCT
    eKind : E_RetainedKind;
    nStation : USINT;               // 0 = machine
    nMover : USINT;
    nId : UDINT;                    // variable, objet ou calibration
    aValue : ARRAY[1..3] OF LREAL;  // valeur ; compteurs : actions, erreurs, heures ; calibration : état
    stPos : ST_Position;
    tStamp : LINT;                  // date de la valeur (calibration)
    sUser : STRING(24);
END_STRUCT
END_TYPE

(* ---- ST_RetainedValues.st ---- *)
// Valeurs rémanentes lues par la HMI (docs/02 § 7.4)
{attribute 'pack_mode' := '1'}
TYPE ST_RetainedValues :
STRUCT
    nRetainId : ULINT;
    nCount : UINT;
    aItem : ARRAY[1..2048] OF ST_RetainedItem;
END_STRUCT
END_TYPE

(* ---- ST_SignalRef.st ---- *)
// Référence vers l'image E/S (docs/04 § 5)
{attribute 'pack_mode' := '1'}
TYPE ST_SignalRef :
STRUCT
    eKind : E_SignalKind;
    nIndex : INT;               // index dans le tableau de GVL_IO correspondant
    bInvert : BOOL;
END_STRUCT
END_TYPE

(* ---- ST_SimForceRequest.st ---- *)
// Forcer une entrée d'un objet simulé (docs/04 § 6.3), Maintenance
{attribute 'pack_mode' := '1'}
TYPE ST_SimForceRequest :
STRUCT
    nSeq : UDINT;
    nStation : USINT;
    nObject : UINT;
    nSignal : USINT;                // S1..S8
    fValue : LREAL;
    bRelease : BOOL;                // faux = forcer, vrai = rendre la main à la simulation
END_STRUCT
END_TYPE

(* ---- ST_SlotStatus.st ---- *)
// Emplacement d'un mover, publié (docs/06 § 6.3)
{attribute 'pack_mode' := '1'}
TYPE ST_SlotStatus :
STRUCT
    bPresent : BOOL;
    sPartId : STRING(40);
    eStatus : E_PartStatus;
    eVerdict : E_Verdict;
    nOrder : UDINT;
END_STRUCT
END_TYPE

(* ---- ST_Staging.st ---- *)
// Zone d'attente du déploiement (docs/06 § 6.2)
{attribute 'pack_mode' := '1'}
TYPE ST_Staging :
STRUCT
    stMachine : ST_MachineData;
    aStation : ARRAY[1..GVL_Const.MAX_STATIONS] OF ST_StationData;
    aPressRecipe : ARRAY[1..GVL_Const.MAX_PRESS_RECIPES] OF ST_PressRecipe;
END_STRUCT
END_TYPE

(* ---- ST_StationCfg.st ---- *)
// Station dans la configuration machine (docs/06 § 4)
{attribute 'pack_mode' := '1'}
TYPE ST_StationCfg :
STRUCT
    bUsed : BOOL;
    sName : STRING(40);
    nGroupMask : UINT;          // bit n-1 = fonction n
    nWorkPos : INT;             // index dans aPlanarPos
    aQueuePos : ARRAY[1..GVL_Const.MAX_QUEUE] OF INT;   // 0 = absente
    fOverride : LREAL;
END_STRUCT
END_TYPE

(* ---- ST_StationData.st ---- *)
// Données déployées d'une station (docs/06 § 4)
{attribute 'pack_mode' := '1'}
TYPE ST_StationData :
STRUCT
    nObjCount : UINT;
    aObj : ARRAY[1..GVL_Const.MAX_OBJ_PER_STATION] OF ST_ObjConfig;   // parents avant enfants
    aTable : ARRAY[1..GVL_Const.MAX_TABLES] OF ST_TableDir;
    nInstrCount : INT;
    aInstr : ARRAY[1..GVL_Const.MAX_INSTR] OF ST_Instr;
    aCond : ARRAY[1..GVL_Const.MAX_COND] OF ST_Condition;
    aText : ARRAY[1..GVL_Const.MAX_TEXTS] OF STRING(80);
    aPos : ARRAY[1..GVL_Const.MAX_NAMED_POS] OF ST_NamedPos;
    aVar : ARRAY[1..GVL_Const.MAX_VARS] OF ST_VarInit;
    aInterlock : ARRAY[1..GVL_Const.MAX_INTERLOCKS] OF ST_Interlock;
    nOpMapCount : USINT;
    aOpMap : ARRAY[1..GVL_Const.MAX_OPMAP] OF ST_OpMap;
    nCalibCount : USINT;
    aCalib : ARRAY[1..GVL_Const.CALIB_PER_STATION] OF ST_CalibDef;
END_STRUCT
END_TYPE

(* ---- ST_StationForce.st ---- *)
// Forçage d'une station (docs/12 § 3)
{attribute 'pack_mode' := '1'}
TYPE ST_StationForce :
STRUCT
    bOutOfProduction : BOOL;
    nReason : USINT;
    tSince : LINT;
    sBy : STRING(24);
END_STRUCT
END_TYPE

(* ---- ST_StationStatus.st ---- *)
// Statut d'une station (docs/06 § 6.3)
{attribute 'pack_mode' := '1'}
TYPE ST_StationStatus :
STRUCT
    eState : E_State;
    eMode : E_Mode;
    fEffOverride : REAL;
    nBeacon : UINT;                 // voir F_BeaconBits
    bFault : BOOL;
    bOutOfProduction : BOOL;
    bQualityLock : BOOL;
    nOpGroup : USINT;
    nOpOperation : USINT;
    nOpMover : USINT;
    nOpSlot : USINT;
    eOpStatus : E_OpStatus;
    fOpElapsedMs : REAL;
    aCtx : ARRAY[1..GVL_Const.MAX_CTX] OF ST_CtxStatus;
    bStepEnabled : BOOL;
    eStepGranularity : E_StepGranularity;
    nCalib : USINT;
    aCalib : ARRAY[1..GVL_Const.CALIB_PER_STATION] OF ST_CalibStatus;
    stPrompt : ST_PromptState;
    nCycleCount : UDINT;
    fLastCycleMs : REAL;
END_STRUCT
END_TYPE

(* ---- ST_StepControl.st ---- *)
// Pas à pas d'une station (docs/05 § 8)
{attribute 'pack_mode' := '1'}
TYPE ST_StepControl :
STRUCT
    bEnabled : BOOL;
    eGranularity : E_StepGranularity;
    nStepSeq : UDINT;               // la HMI l'incrémente pour autoriser un pas
END_STRUCT
END_TYPE

(* ---- ST_TableDir.st ---- *)
// Répertoire des tables (docs/06 § 2)
{attribute 'pack_mode' := '1'}
TYPE ST_TableDir :
STRUCT
    bUsed : BOOL;
    sName : STRING(40);
    eKind : E_TableKind;
    nStart : INT;               // index de la première instruction dans aInstr
    nLength : INT;
END_STRUCT
END_TYPE

(* ---- ST_TraceBuffer.st ---- *)
// Tampon de traces (docs/05 § 9)
{attribute 'pack_mode' := '1'}
TYPE ST_TraceBuffer :
STRUCT
    nWriteSeq : UDINT;
    aTrace : ARRAY[0..GVL_Const.TRACE_BUFFER - 1] OF ST_TraceRecord;
END_STRUCT
END_TYPE

(* ---- ST_TraceRecord.st ---- *)
// Trace d'une opération sur une pièce (docs/05 § 9)
{attribute 'pack_mode' := '1'}
TYPE ST_TraceRecord :
STRUCT
    nSeq : UDINT;
    sPartId : STRING(40);
    nOrder : UDINT;
    nMover : USINT;
    nSlot : USINT;
    nStation : USINT;
    nGroup : USINT;
    nOperation : USINT;
    tStart : LINT;
    tEnd : LINT;
    eVerdict : E_Verdict;
    nErrorCode : UINT;
    aData : ARRAY[1..GVL_Const.MAX_PART_DATA] OF LREAL;
    nCurveId : UDINT;               // 0 = aucune
END_STRUCT
END_TYPE

(* ---- ST_Value.st ---- *)
// Valeur d'un paramètre d'instruction (docs/06 § 2), 11 octets
{attribute 'pack_mode' := '1'}
TYPE ST_Value :
STRUCT
    eSource : E_ValueSource;
    nIndex : INT;               // n° de variable, donnée, paramètre, position, vitesse, texte, objet, variable système
    fValue : LREAL;             // constante ; ObjValue : n° de valeur E1..E4 ; position : décalage ajouté
END_STRUCT
END_TYPE

(* ---- ST_VarInit.st ---- *)
// Déclaration d'une variable de station (docs/06 § 2)
{attribute 'pack_mode' := '1'}
TYPE ST_VarInit :
STRUCT
    eType : E_VarType;
    fValue : LREAL;
    stPos : ST_Position;
    bRetain : BOOL;             // persistante (calibration), conservée au redéploiement par identifiant
    nId : UDINT;                // identifiant stable (empreinte de l'Id du projet) ; 0 = variable cachée (D92)
END_STRUCT
END_TYPE
